TYPE st_TankValves :
STRUCT
	valOutlet		: E_Pis_Name;//Comment?
	valLine			: E_Pis_Name;//Comment?
	valTriBlender	: E_Pis_Name;//Comment?
	valDrain		: E_Pis_Name;//Comment?
	valCIP			: E_Pis_Name;//Comment?
END_STRUCT
END_TYPE

(* stored: Version 1.1.0.1, ProductVersion 3.1.4024.12
   DUT st_TankValves: Id {ef0ebba3-3648-41a3-8037-3a8b29bb75df} *)
